Fanuc KAREL source: kf00038.KL

-- PROVISIONAL review KL for V770-1; original PC SHA256 213de98af7c221fbd0ccaec4581120b8307b20e9dbb8337117d037453aa9132a
-- Incomplete behavior may be omitted. Consult companion uncertainty JSON. Do not deploy.
PROGRAM KF00038
%NOLOCKGROUP
VAR
  I : INTEGER
  J : INTEGER
  X : REAL
  Y : REAL
  B : BOOLEAN
  C : BOOLEAN
  TXT : STRING[80]
  TXT2 : STRING[80]
  STATUS : INTEGER
-- UNRESOLVED_DECL AI type=002010
-- UNRESOLVED_DECL BI type=002010
-- UNRESOLVED_DECL P type=000102
-- UNRESOLVED_DECL JP type=000199
-- UNRESOLVED_DECL PF type=000101
-- UNRESOLVED_DECL V1 type=000013
-- UNRESOLVED_DECL V2 type=000013
BEGIN
  -- UNRESOLVED_PC offsets 5-19; opcodes 2E,22,9D,33,35
  -- UNRESOLVED_PC offsets 24-38; opcodes 22,22,1E
  -- UNRESOLVED_PC offsets 43-47; opcodes 7F
END KF00038
